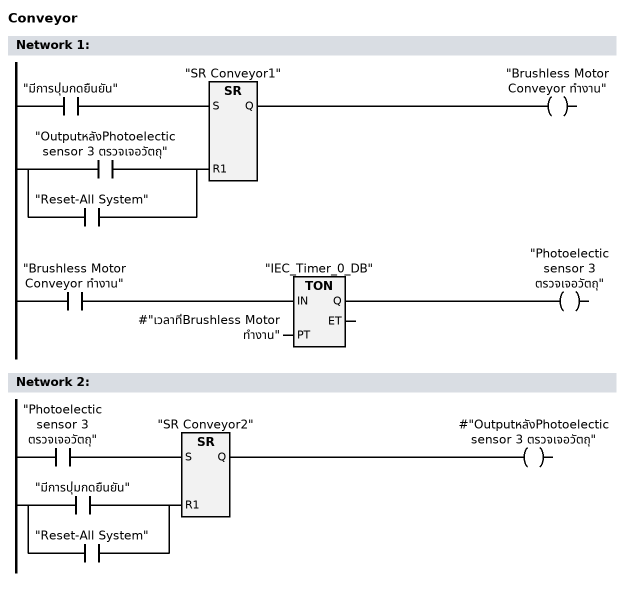
   IF "มีการปุ่มกดยืนยัน" THEN
       "SR Conveyor1" := TRUE;   // SR flip-flop
   END_IF;
   IF "OutputหลังPhotoelectic sensor 3 ตรวจเจอวัตถุ" OR "Reset-All System" THEN
       "SR Conveyor1" := FALSE;
   END_IF;
   "Brushless Motor Conveyor ทำงาน" := "SR Conveyor1";
   "IEC_Timer_0_DB".TON(IN := "Brushless Motor Conveyor ทำงาน", PT := #"เวลาที่Brushless Motor ทำงาน");
   "Photoelectic sensor 3 ตรวจเจอวัตถุ" := "IEC_Timer_0_DB".Q;
END_REGION

REGION Network 2
   RUNG wire#powerrail
      Contact( "Photoelectic sensor 3 ตรวจเจอวัตถุ" )
      S_SR(operand := "SR Conveyor2", r1 := wire#w1)
      Coil( #"OutputหลังPhotoelectic sensor 3 ตรวจเจอวัตถุ" )
   END_RUNG
   RUNG wire#powerrail
      Contact( "มีการปุ่มกดยืนยัน" )
   END_RUNG wire#w1
   RUNG wire#powerrail
      Contact( "Reset-All System" )
   END_RUNG wire#w1
   // the same network as SCL:
   IF "Photoelectic sensor 3 ตรวจเจอวัตถุ" THEN
       "SR Conveyor2" := TRUE;   // SR flip-flop
   END_IF;
   IF "มีการปุ่มกดยืนยัน" OR "Reset-All System" THEN "SR Conveyor2" := FALSE; END_IF;
   #"OutputหลังPhotoelectic sensor 3 ตรวจเจอวัตถุ" := "SR Conveyor2";
END_REGION
END_FUNCTION

// folder: System_In(จัดเก็บ)

FUNCTION "Memory_Bacode" : Void   // FC2, LAD
{ S7_Optimized_Access := 'TRUE' }
VERSION : 0.1
   VAR_OUTPUT
      "Output Barcode" : Bool;
   END_VAR
BEGIN

REGION Network 1
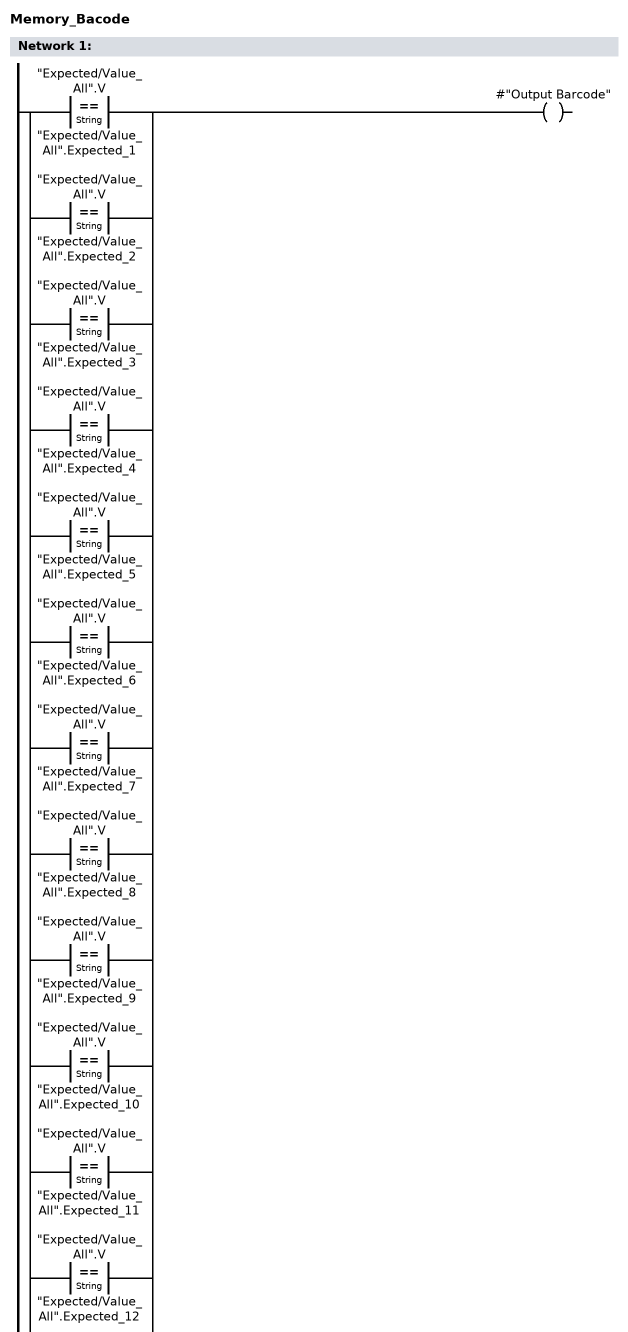
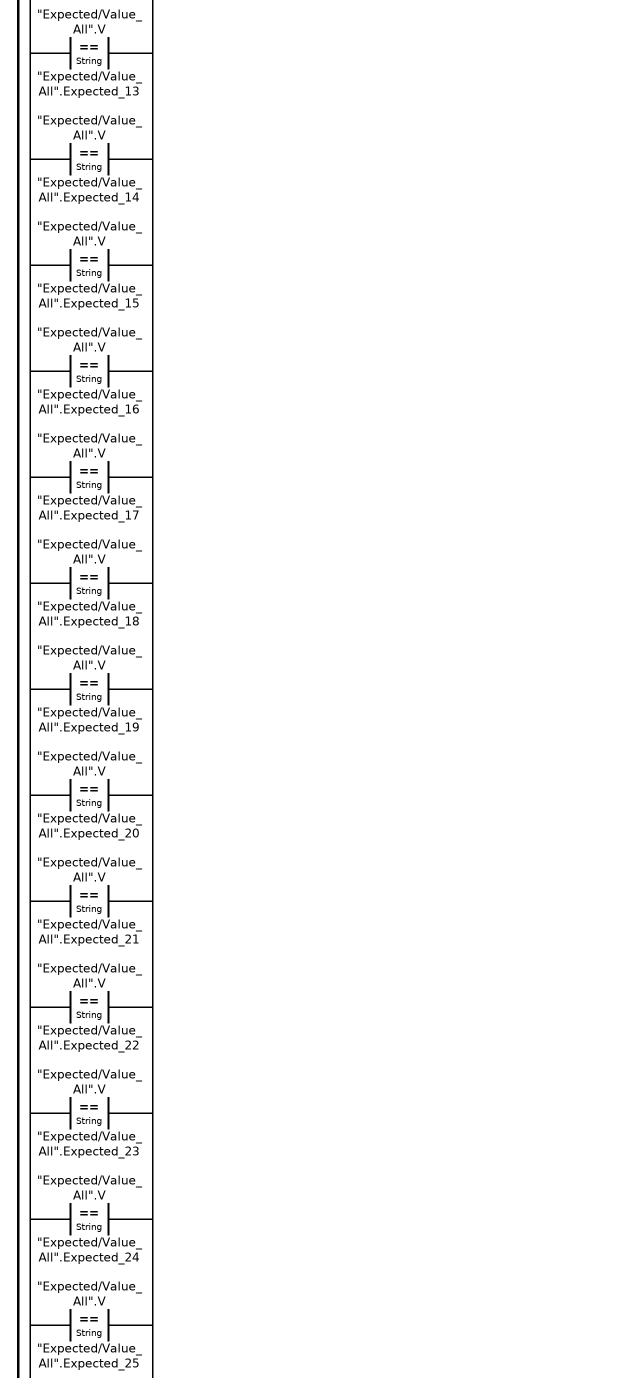
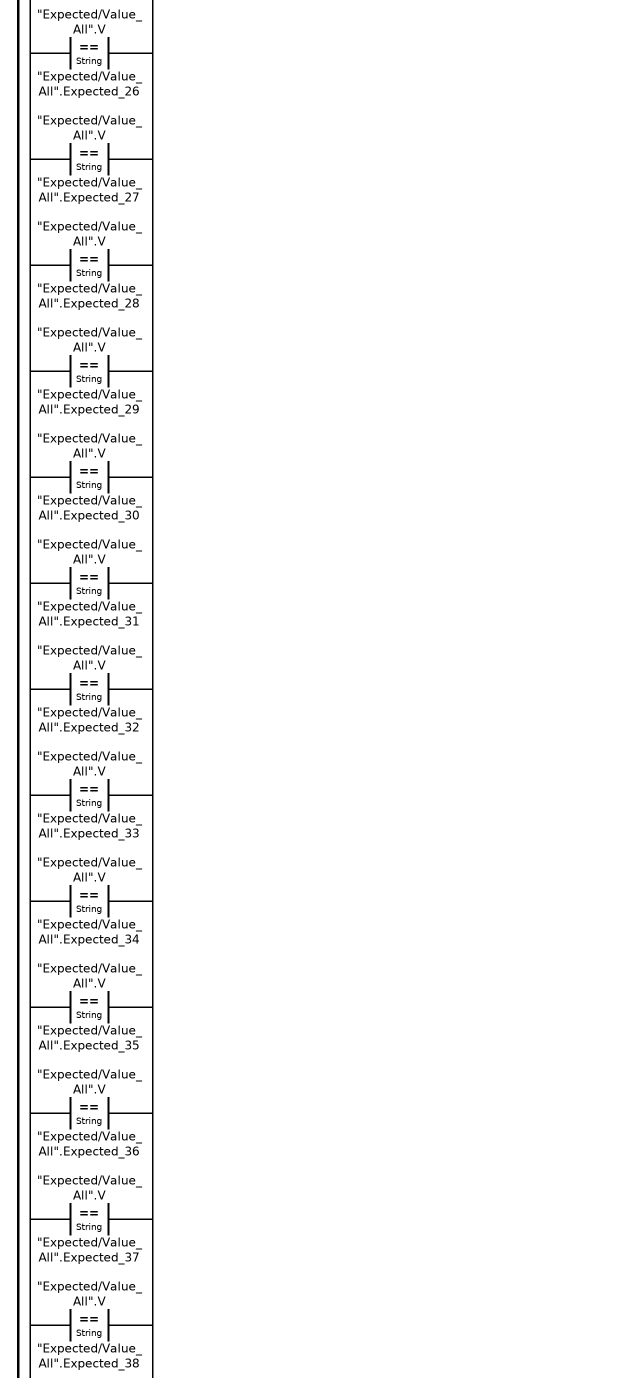
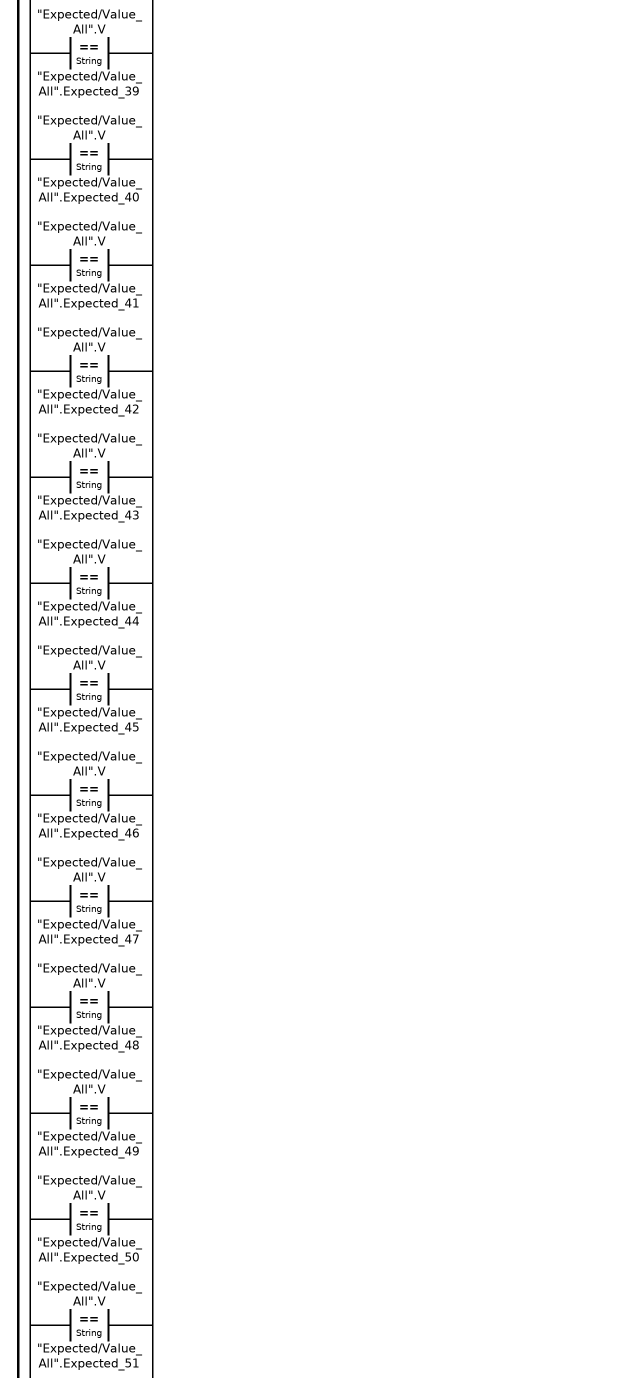
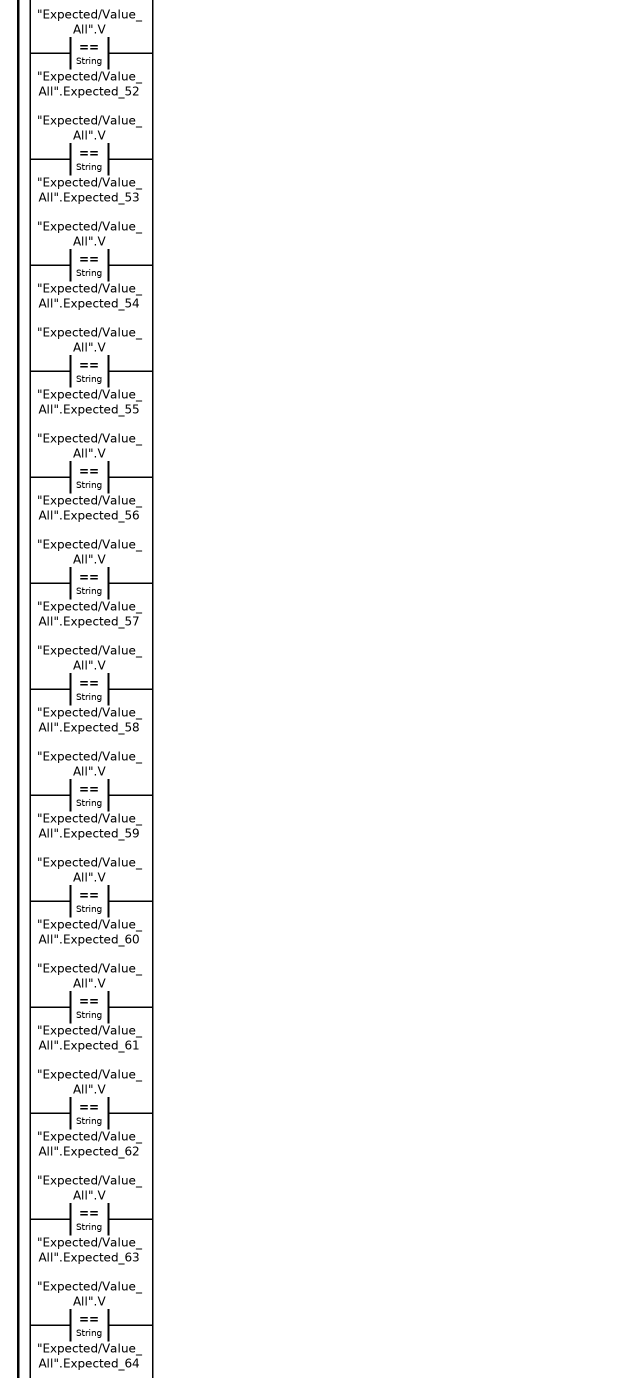
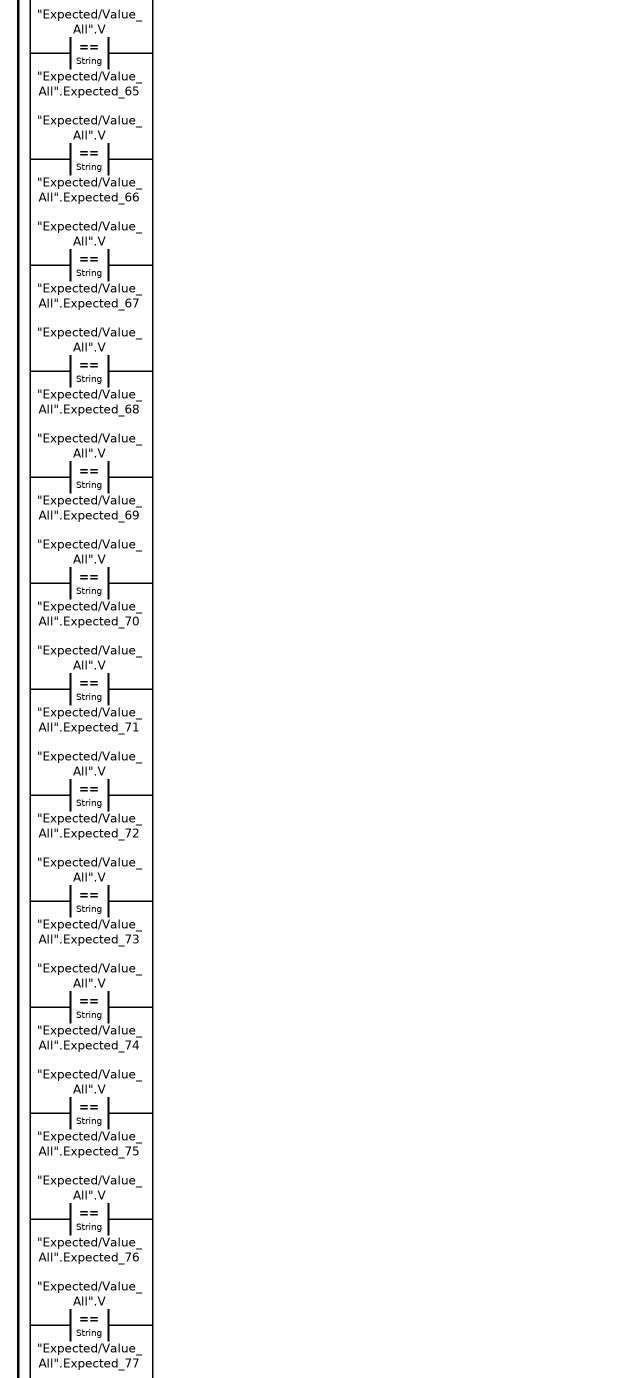
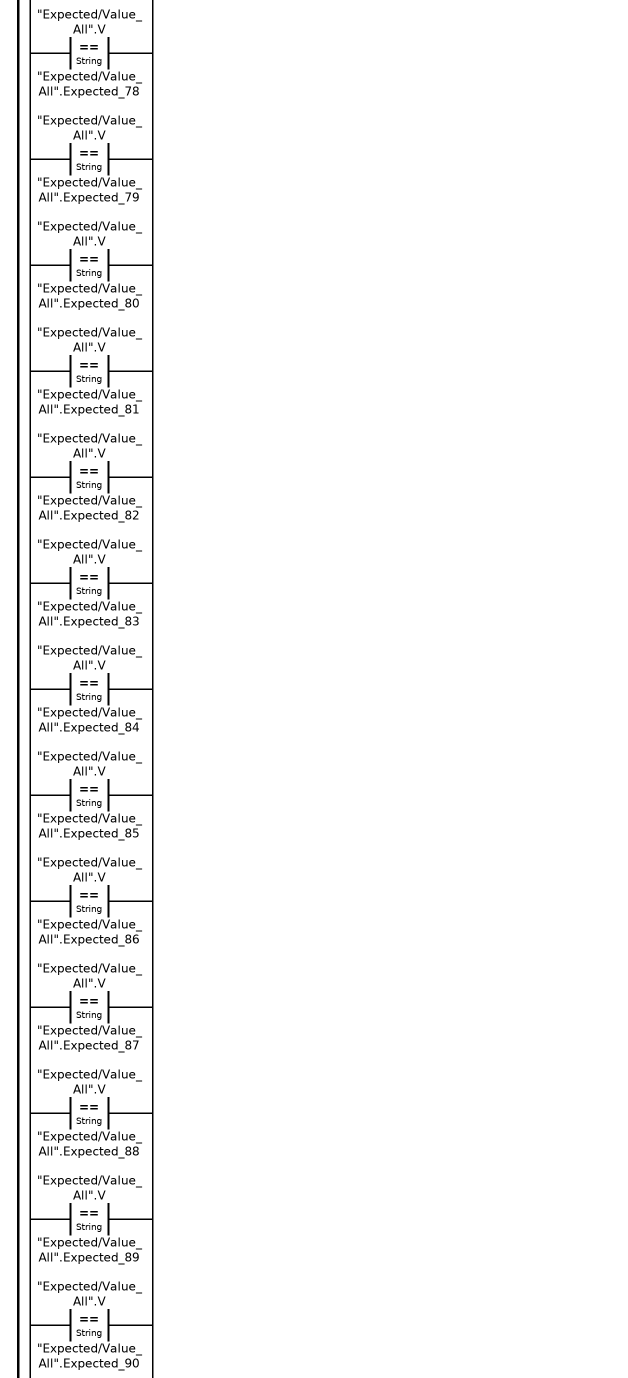
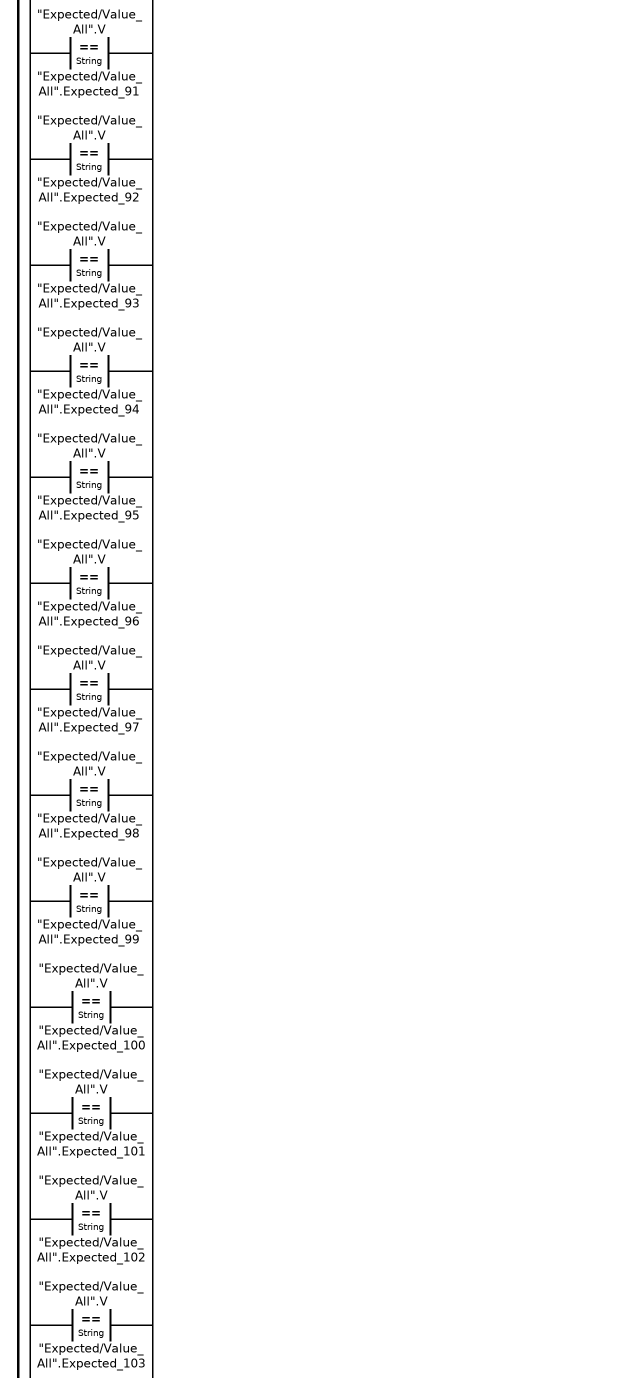
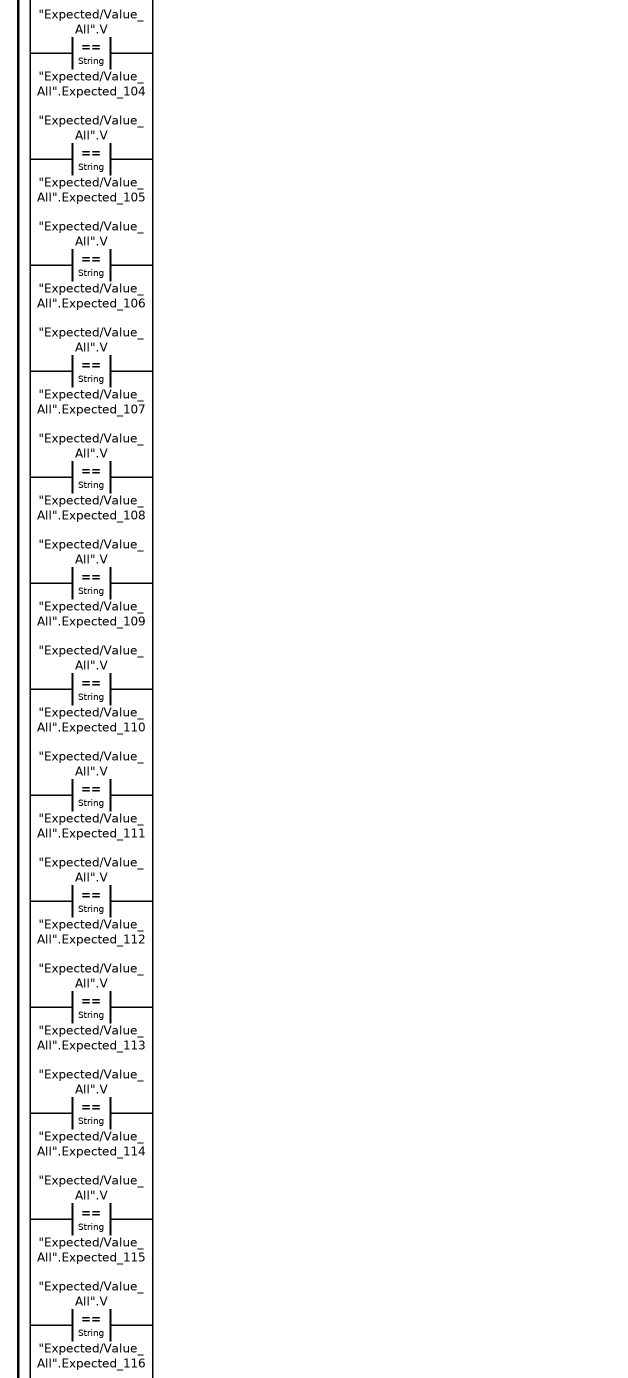
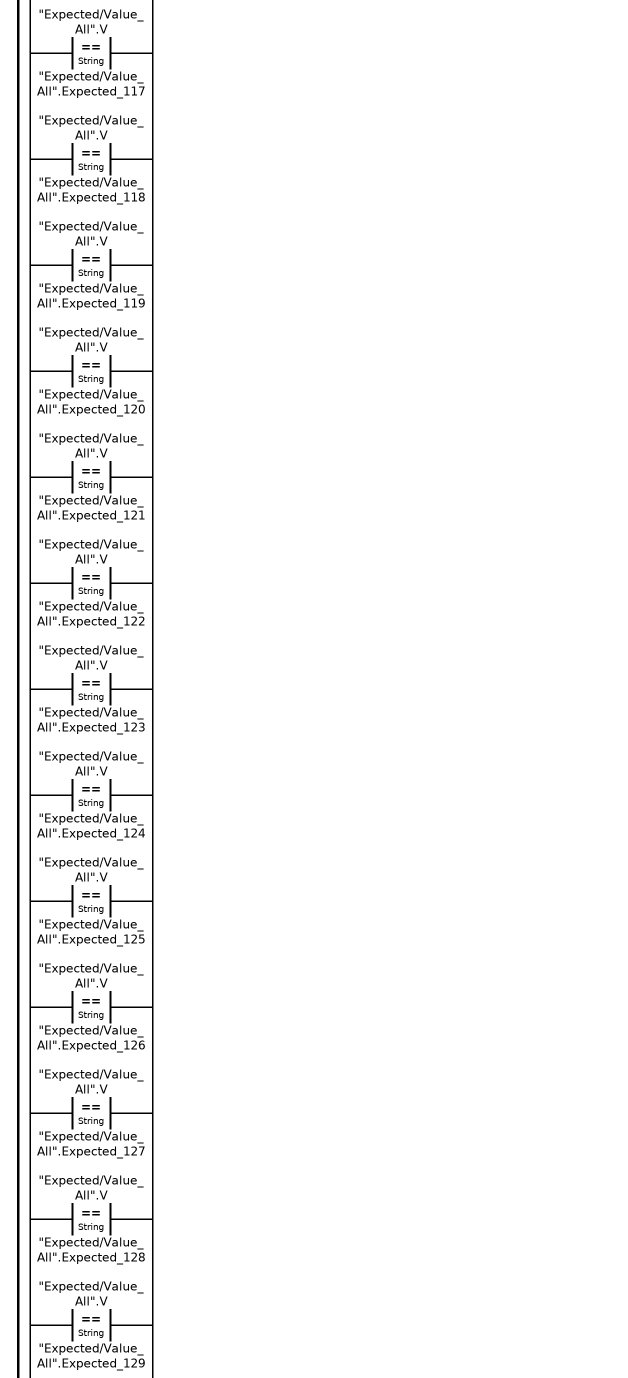
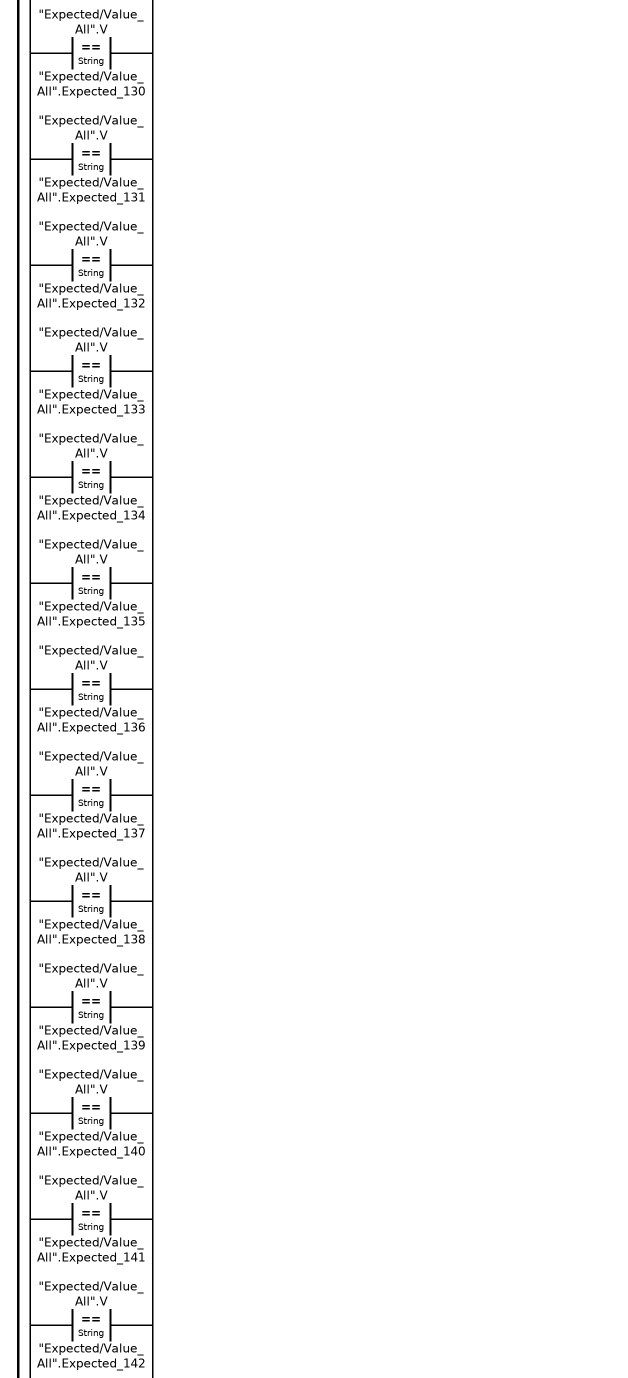
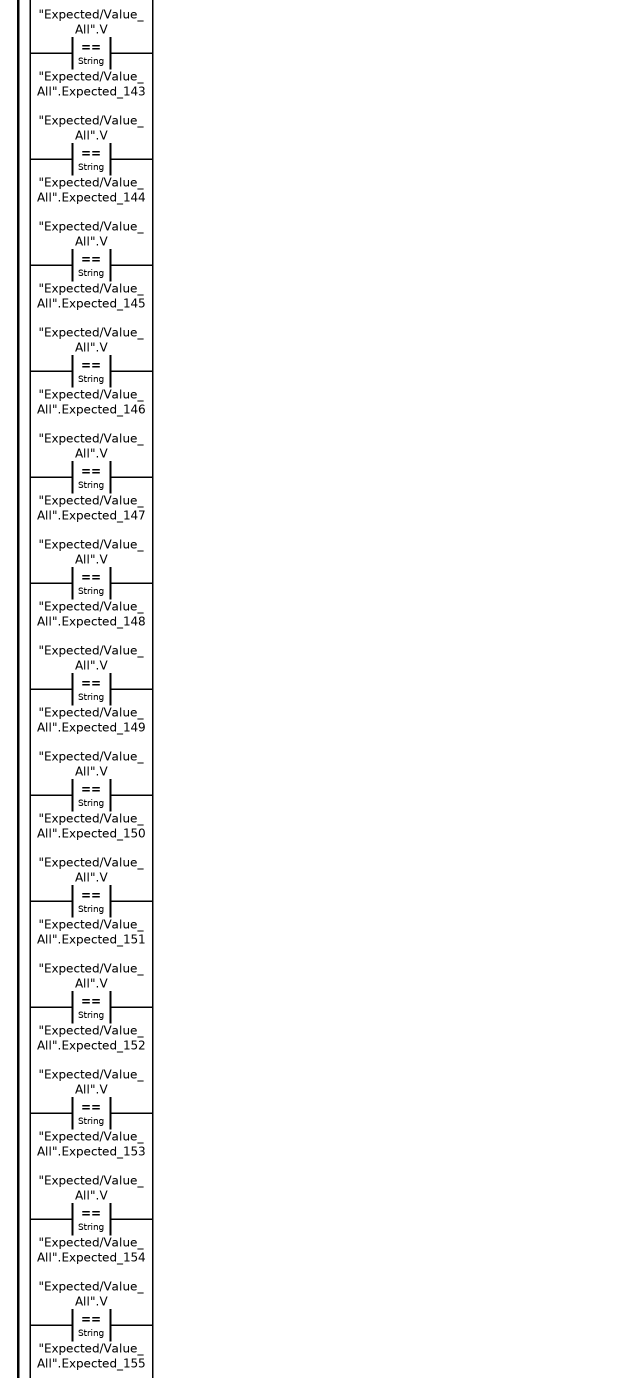
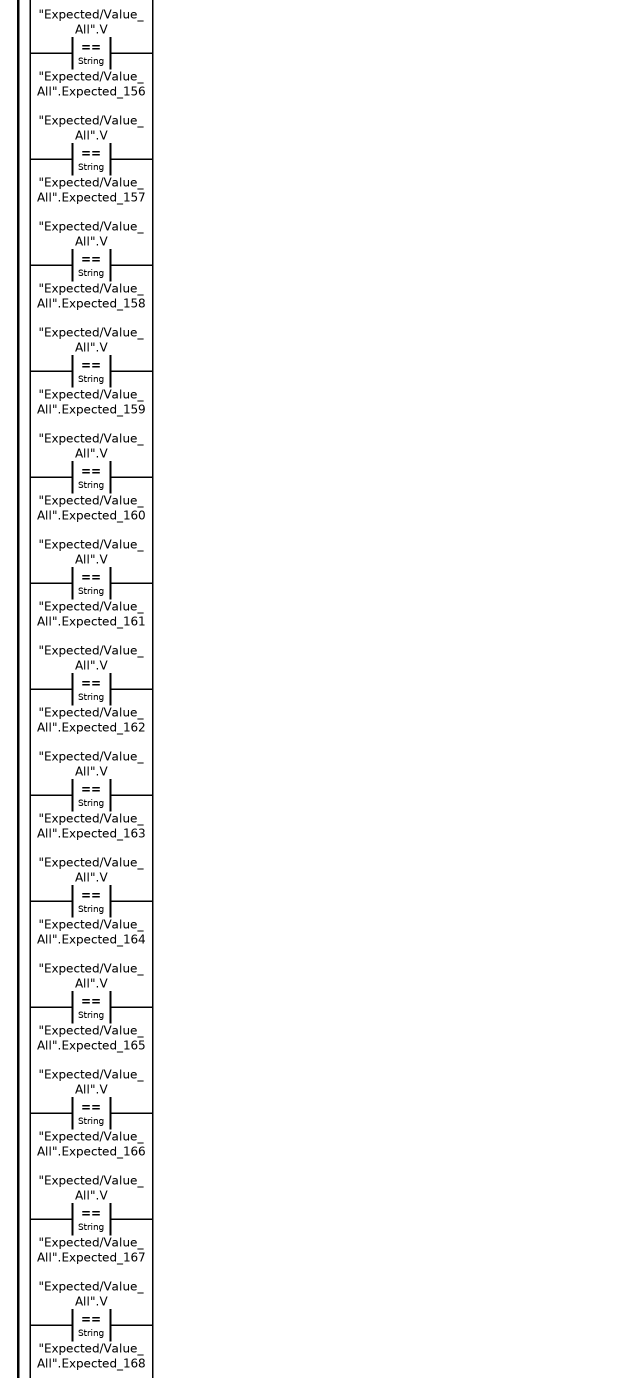
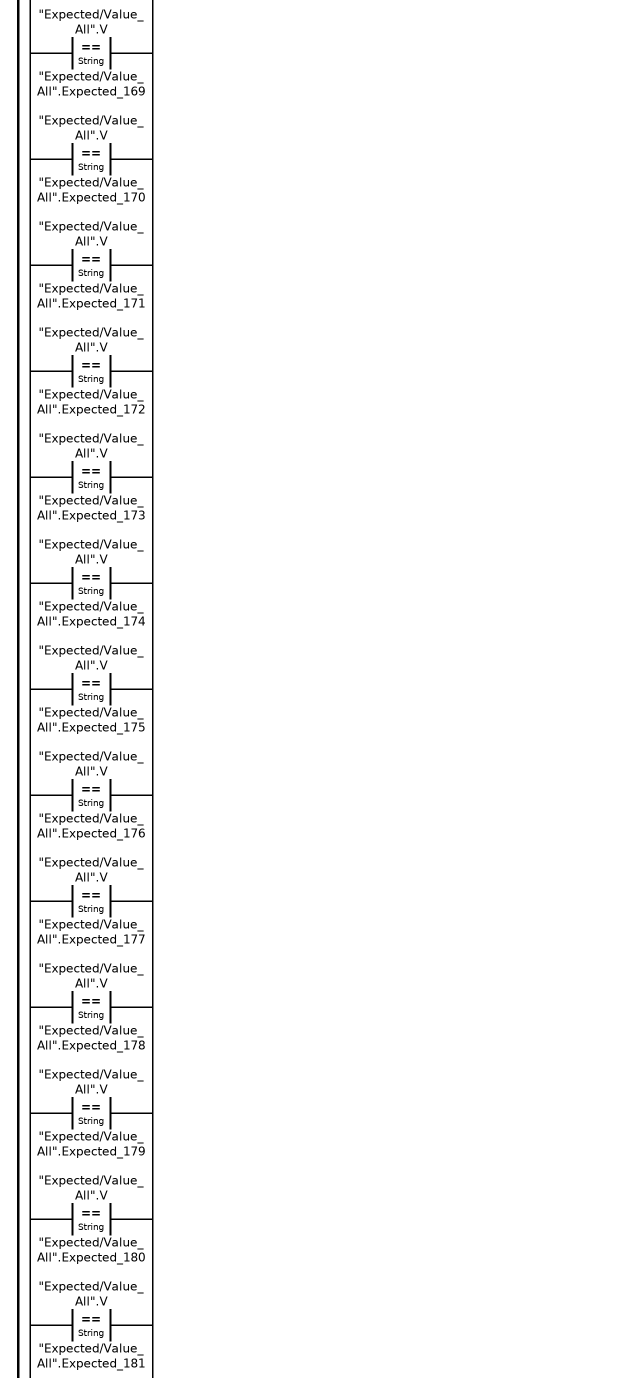
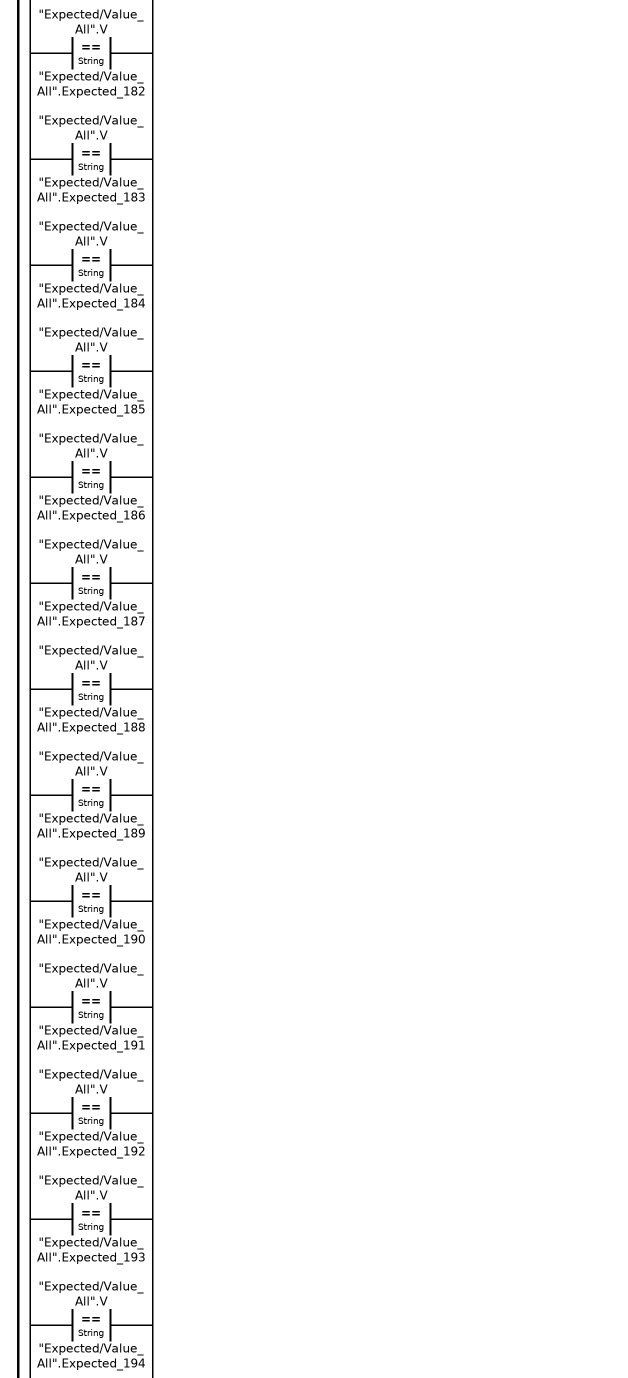
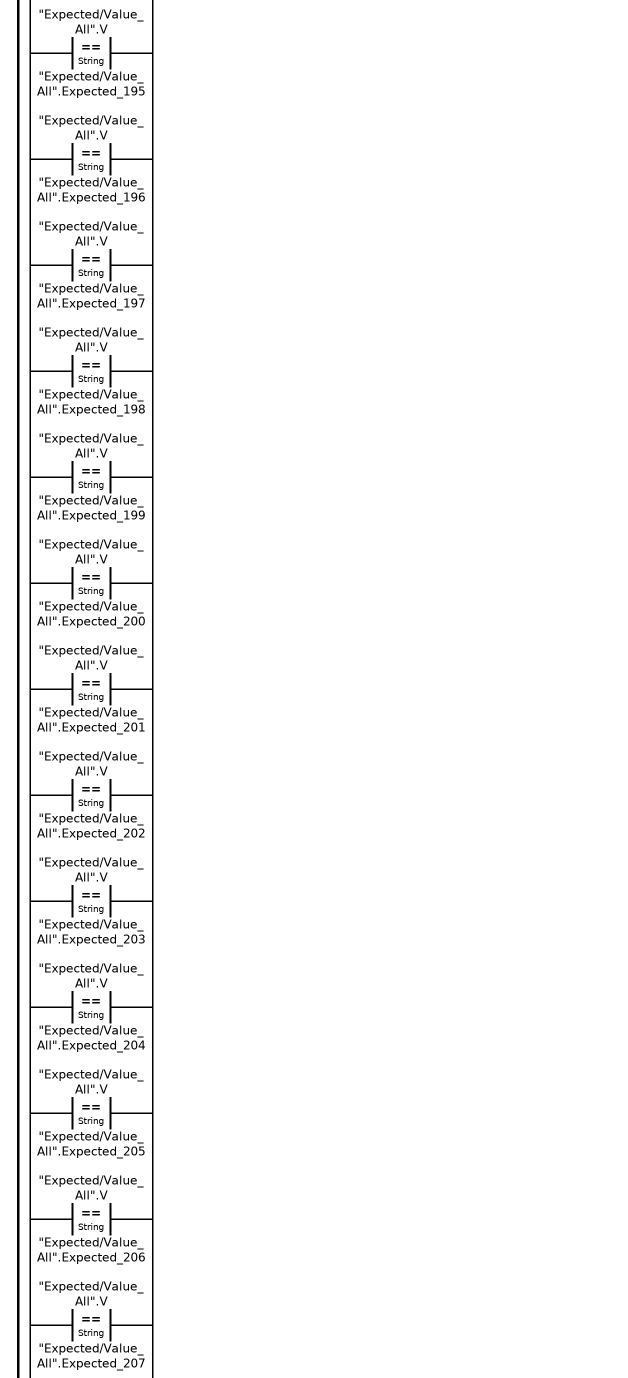
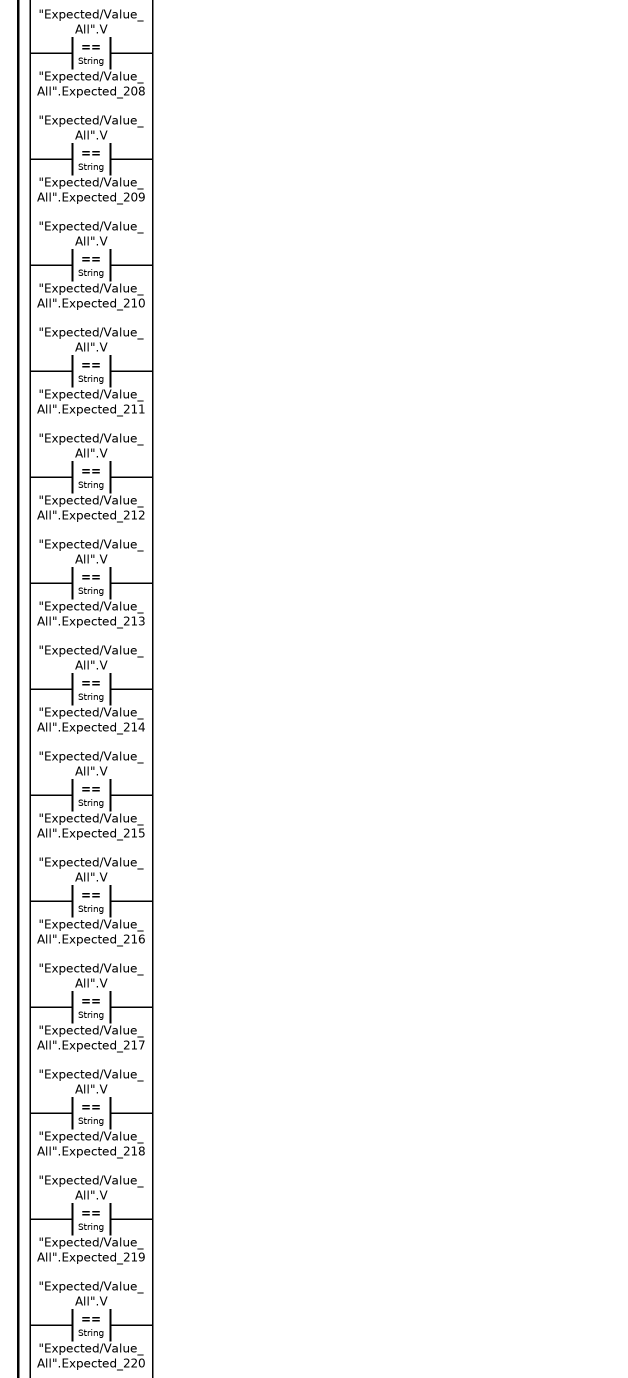
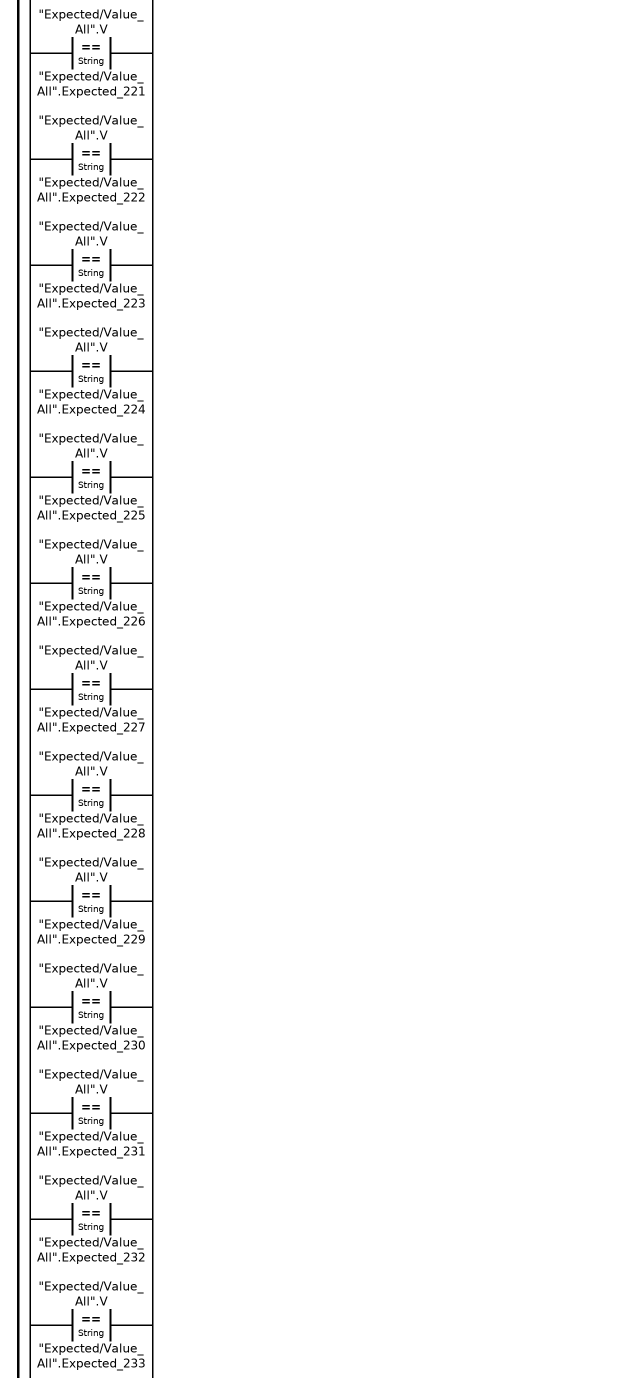
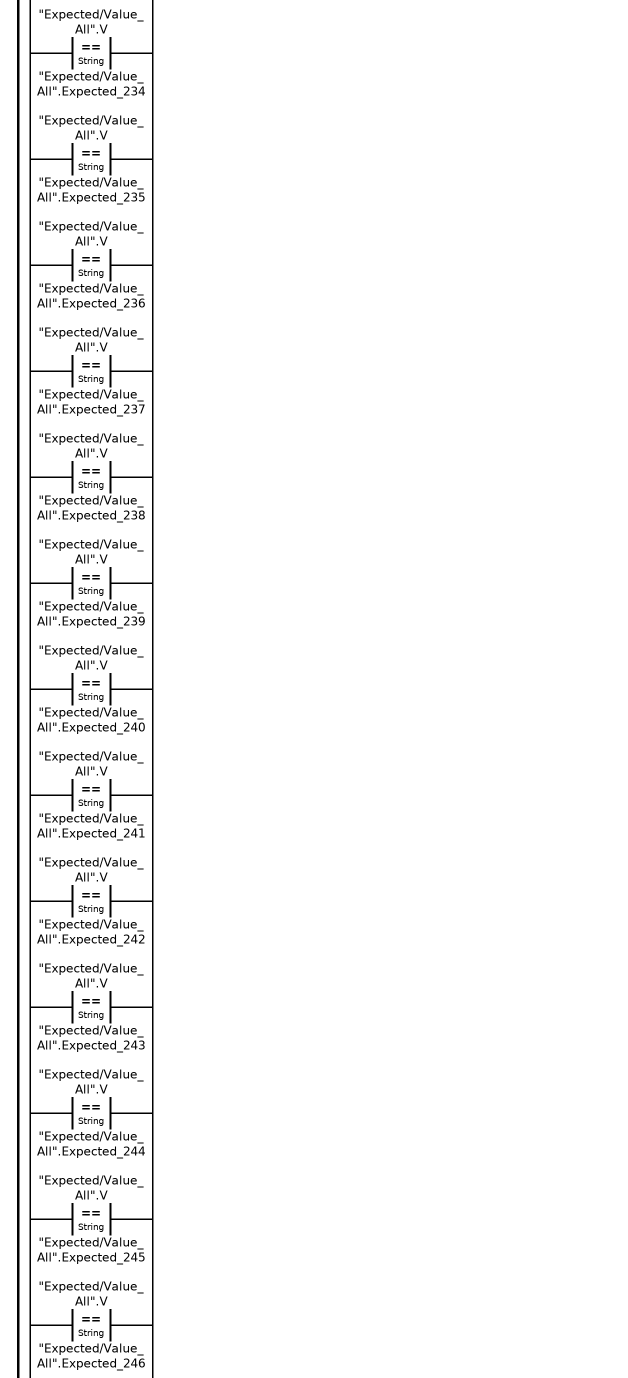
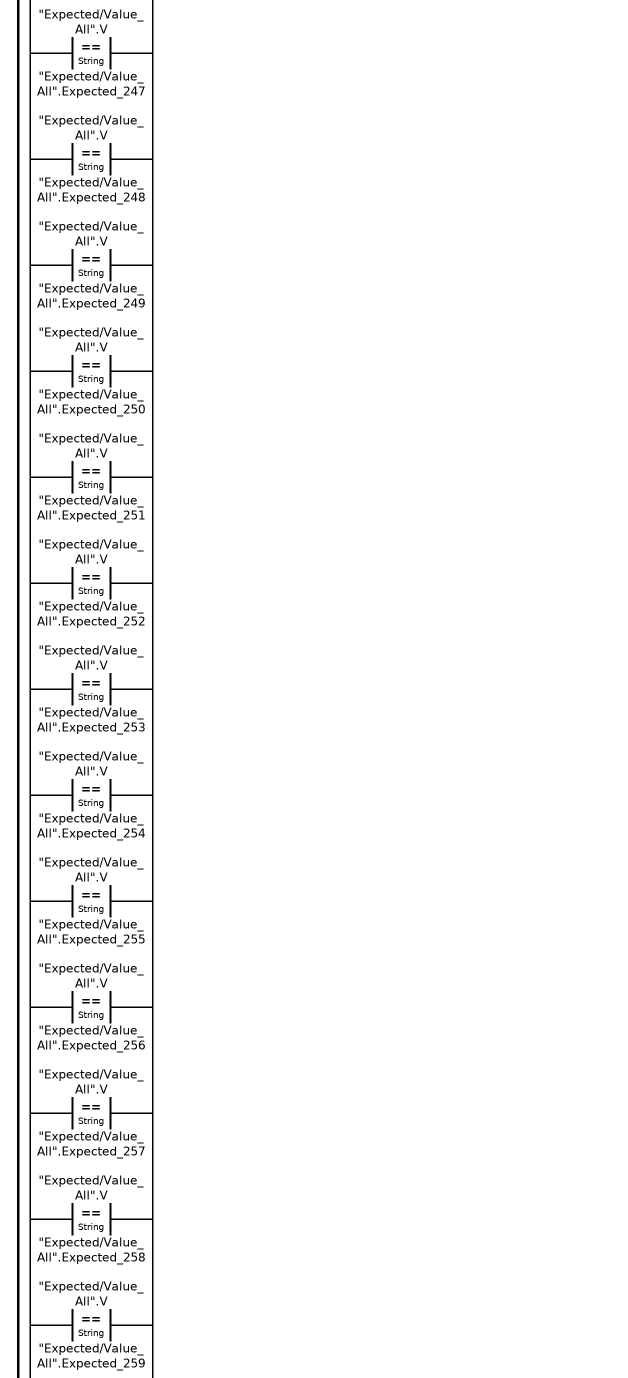
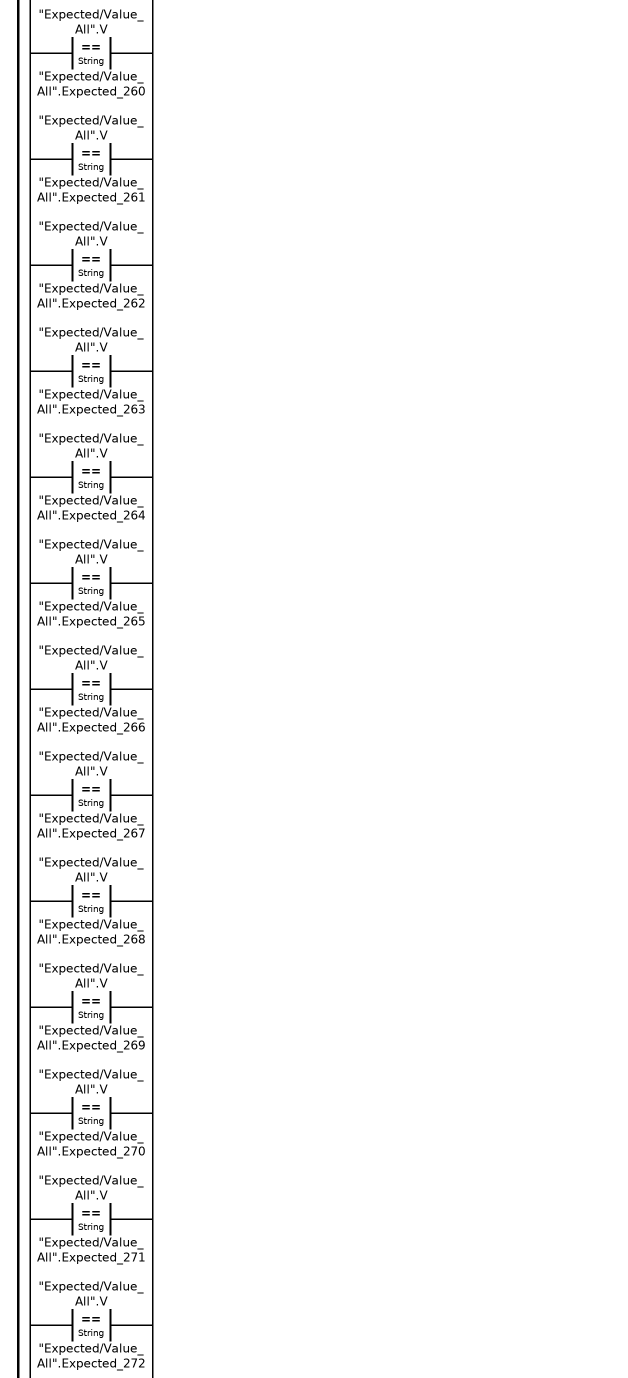
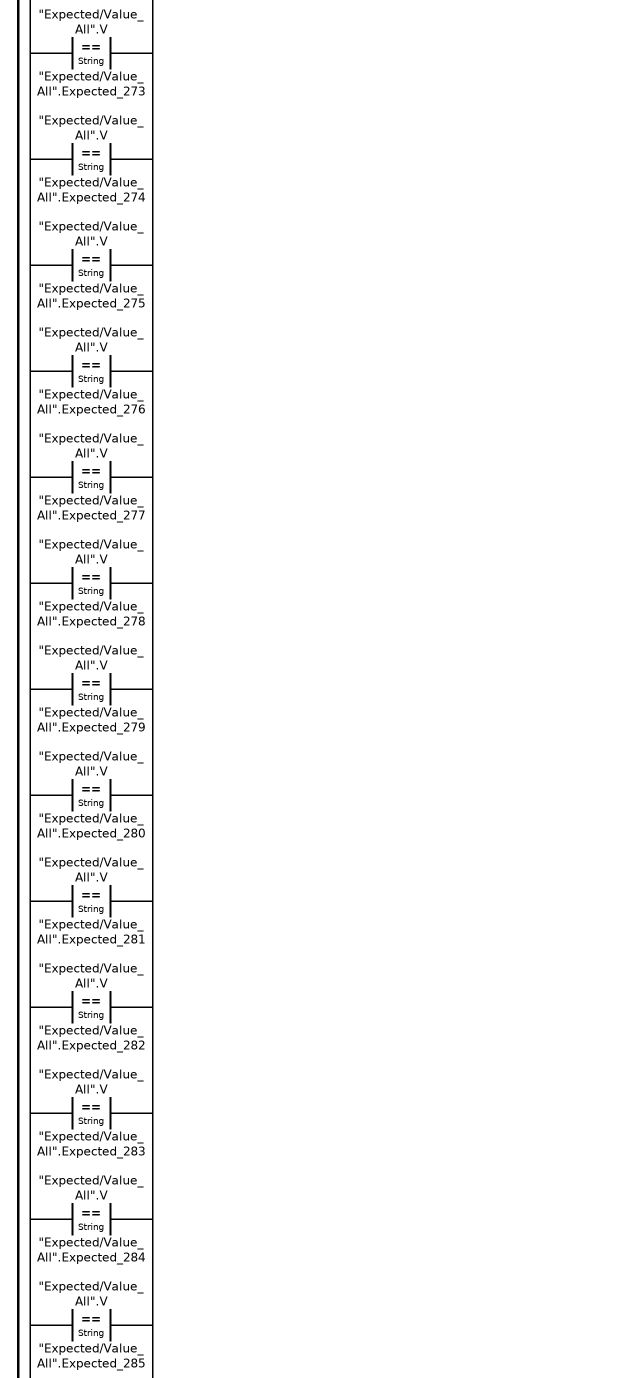
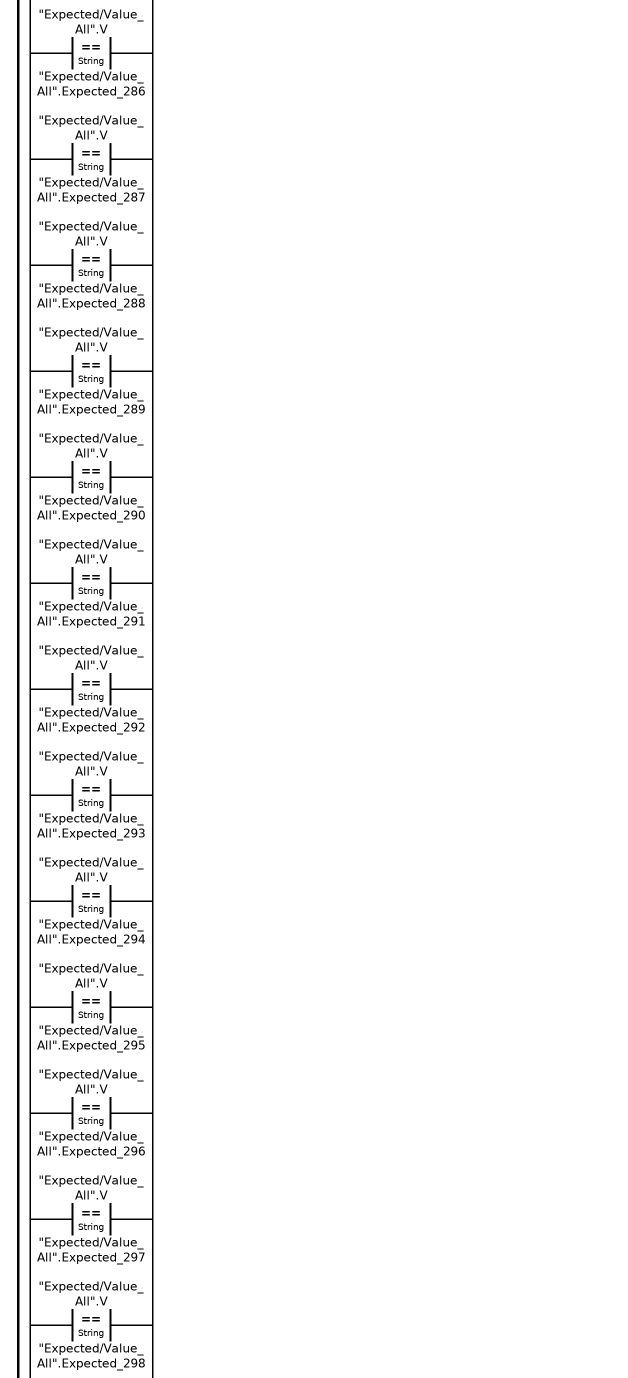
